Staubli VAL3: utCommon.dtx

public string sText
public string sID
public string sPage
